// Generated by voz_llm_plc_agent
// Target: Siemens TIA Portal V18 - SCL external source
// Review and compile before any download to physical hardware.

FUNCTION_BLOCK "PLC_PRG"
{ S7_Optimized_Access := 'TRUE' }
VERSION : 0.1
VAR_INPUT
   I_Emergency : Bool := FALSE;
   I_Start : Bool := FALSE;
END_VAR
VAR_OUTPUT
   Q_Motor_Enable : Bool := FALSE;
END_VAR
VAR
   M_Cond1_Prev : Bool;
   M_Cond1_Active : Bool;
   T_Cond1 {InstructionName := 'TON_TIME'; LibVersion := '1.0'} : TON_TIME;
END_VAR
BEGIN
(* Salida condicionada 1: pulso de T#3s al cumplirse la condicion *)
IF (#I_Start AND NOT #I_Emergency) AND NOT #M_Cond1_Prev THEN
    #M_Cond1_Active := TRUE;
END_IF;
#M_Cond1_Prev := (#I_Start AND NOT #I_Emergency);
#T_Cond1(IN := #M_Cond1_Active, PT := T#3s);
IF #T_Cond1.Q THEN
    #M_Cond1_Active := FALSE;
END_IF;
(* Salidas: contribucion automatica (secuencia/condiciones) y manual, con sus bloqueos *)
#Q_Motor_Enable := #M_Cond1_Active AND NOT #I_Emergency;
END_FUNCTION_BLOCK

DATA_BLOCK "DB_PLC_PRG"
{ S7_Optimized_Access := 'TRUE' }
VERSION : 0.1
NON_RETAIN
"PLC_PRG"
BEGIN
END_DATA_BLOCK

ORGANIZATION_BLOCK "Main"
{ S7_Optimized_Access := 'TRUE' }
VERSION : 0.1
BEGIN
   "DB_PLC_PRG"(
      I_Emergency := "I_Emergency",
      I_Start := "I_Start",
      Q_Motor_Enable => "Q_Motor_Enable"
   );
END_ORGANIZATION_BLOCK
